(* IEC 61131-3 sources: STAR-PLC-Agent/results/raw/codex_terra_pilot_20261114/PUB001/formal/attempt_0001, 1 file *)

(* ---- candidate.st ---- *)
FUNCTION_BLOCK FB_Task
VAR_INPUT
    bottleSensor : BOOL;
    cleaningConfirmButton : BOOL;
    fillingConfirmButton : BOOL;
    cappingConfirmButton : BOOL;
    packingConfirmButton : BOOL;
    finishedButton : BOOL;
END_VAR
VAR_OUTPUT
    Pump_Motor : BOOL := FALSE;
    Filling_Valve : BOOL := FALSE;
    Capping_Machine : BOOL := FALSE;
    Packing_Machine : BOOL := FALSE;
    Completion_Light : BOOL := FALSE;
END_VAR
VAR
    phase : INT := 0;
END_VAR

CASE phase OF
    0:
        IF bottleSensor THEN
            phase := 1;
        END_IF;
    1:
        IF cleaningConfirmButton THEN
            phase := 2;
        END_IF;
    2:
        IF fillingConfirmButton THEN
            phase := 3;
        END_IF;
    3:
        IF cappingConfirmButton THEN
            phase := 4;
        END_IF;
    4:
        IF packingConfirmButton THEN
            phase := 5;
        END_IF;
    5:
        IF finishedButton THEN
            phase := 0;
        END_IF;
END_CASE;

Pump_Motor := phase = 1;
Filling_Valve := phase = 2;
Capping_Machine := phase = 3;
Packing_Machine := phase = 4;
Completion_Light := phase = 5;
END_FUNCTION_BLOCK
